(* IEC 61131-3 sources: nautilus/logix/deploy/testdata, 1 file *)

(* ---- keep_types.st ---- *)
TYPE
  LineStatus : STRUCT
    Mode  : DINT;
    Alarm : BOOL;
  END_STRUCT;
  Pump : STRUCT
    Run    : BOOL;
    Speed  : REAL;
    Status : LineStatus;
  END_STRUCT;
END_TYPE
